Fanuc KAREL source: KT00709.KL

PROGRAM KT00709
%NOLOCKGROUP
VAR
  R1: REAL
  R2: REAL
  OUT: INTEGER
BEGIN
  R1 = 2.0
  R2 = 3.0
  R1 = 2.0
  R2 = 3.0
  OUT = ARRAY_LEN(R1)
END KT00709
